{attribute 'linkalways'}
{attribute 'no_explicit_call' := 'This FB is a CLASS and must be accessed using methods or properties'}
{attribute 'enable_dynamic_creation'}
FUNCTION_BLOCK Node_F_VN_ConvertDataLayout EXTENDS VisionNode
VAR
    ipSrcImage : _ITcVnImage;
    ipDestImage : _ITcVnImage;
    nSrcDataLayout : _ULINT(ETcVnDataLayout.TCVN_DL_DEFAULT);
    nDestDataLayout : _ULINT(ETcVnDataLayout.TCVN_DL_3D_CHW);
    hrPrev : _HRESULT(S_OK);
    hresult : _HRESULT(S_OK);
END_VAR

METHOD PUBLIC Clone : I_Node
VAR
    pNode : POINTER TO Node_F_VN_ConvertDataLayout;
END_VAR
pNode := __NEW(Node_F_VN_ConvertDataLayout);
Clone := pNode^;
END_METHOD

METHOD FB_init : BOOL
VAR_INPUT
    bInitRetains : BOOL;
    bInCopyCode : BOOL;
END_VAR
AddInput('ipSrcImage', ipSrcImage);
AddParameter('nSrcDataLayout', nSrcDataLayout);
AddParameter('nDestDataLayout', nDestDataLayout);
AddInput('hrPrev', hrPrev);
AddOutput('ipDestImage', ipDestImage);
AddOutput('hresult', hresult);
END_METHOD

METHOD PROTECTED OnExecute
hresult.Value := F_VN_ConvertDataLayout(
    ipSrcImage := ipSrcImage.Value,
    ipDestImage := ipDestImage.Value,
    nSrcDataLayout := nSrcDataLayout.Value,
    nDestDataLayout := nDestDataLayout.Value,
    hrPrev := hrPrev.Value);
END_METHOD

METHOD PUBLIC PreExecutionCheck
VAR_INPUT
    Check : I_PreExecutionChecks;
END_VAR
Check.IsTrue(ipSrcImage.IsValid, 'ipSrcImage must contain an image');
Check.IsTrue((nDestDataLayout.Value <> 0) AND (nDestDataLayout.Value <> ETcVnDataLayout.TCVN_DL_DEFAULT), 'nDestDataLayout must not be 0 or TCVN_DL_DEFAULT');
END_METHOD

END_FUNCTION_BLOCK

(* stored: Version 1.1.0.1, ProductVersion 3.1.4026.19
   POU Node_F_VN_ConvertDataLayout: Id {6df592f4-414e-42ca-bfec-c3d85275f074}, SpecialFunc None
   Folder Constructor: Id {b4d7e482-a8e0-4bb3-841b-4864528fdb6f}
   Method Clone: Id {438af4f9-1988-4d80-9edf-2e61d972ce19}
   Method FB_init: Id {9887a487-9c66-4483-8939-22e2a728266b}
   Method OnExecute: Id {33c2ec74-8c97-4763-8050-3cb08a913c21}
   Method PreExecutionCheck: Id {9cded2d8-3487-4ba3-b139-3149b2ef314d} *)
